FUNCTION_BLOCK FB_ConveyorBase IMPLEMENTS I_Conveyor
VAR_OUTPUT
    initCount : DINT;
    cycleCount : DINT;
END_VAR
VAR
    startup : TON;
    productEdge : R_TRIG;
    delay : TIME;
    requested : BOOL;
    runningState : BOOL;
    lastBlocked : BOOL;
    alarmText : STRING(80);
    count : DINT;
    speed : REAL;
END_VAR

(* All behavior is called through the interface methods. *)

METHOD PUBLIC FB_init : BOOL
VAR_INPUT
    bInitRetains : BOOL;
    bInCopyCode : BOOL;
    startDelay : TIME;
END_VAR
delay := startDelay;
initCount := initCount + 1;
FB_init := TRUE;
END_METHOD

METHOD PUBLIC Start
IF alarmText = '' THEN requested := TRUE; END_IF;
END_METHOD

METHOD PUBLIC Stop
requested := FALSE;
runningState := FALSE;
startup(IN := FALSE, PT := delay);
END_METHOD

METHOD PUBLIC Reset
IF NOT lastBlocked THEN alarmText := ''; END_IF;
END_METHOD

METHOD PROTECTED DetectJam : BOOL
VAR_INPUT
    blocked : BOOL;
END_VAR
DetectJam := FALSE;
END_METHOD

METHOD PUBLIC Cycle
VAR_INPUT
    enabled : BOOL;
    sensor : BOOL;
    blocked : BOOL;
END_VAR
cycleCount := cycleCount + 1;
lastBlocked := blocked;
IF THIS^.DetectJam(blocked := blocked) THEN
    alarmText := 'Jammed';
    requested := FALSE;
END_IF;
startup(IN := requested AND enabled AND alarmText = '', PT := delay);
runningState := startup.Q;
productEdge(CLK := sensor);
IF runningState AND productEdge.Q THEN count := count + 1; END_IF;
END_METHOD

PROPERTY PUBLIC Running : BOOL
GET
Running := runningState;
END_GET
END_PROPERTY

PROPERTY PUBLIC Alarm : STRING(80)
GET
Alarm := alarmText;
END_GET
END_PROPERTY

PROPERTY PUBLIC ProductCount : DINT
GET
ProductCount := count;
END_GET
END_PROPERTY

PROPERTY PUBLIC ActualSpeed : REAL
GET
IF runningState THEN ActualSpeed := speed; ELSE ActualSpeed := 0.0; END_IF;
END_GET
END_PROPERTY

PROPERTY PUBLIC SpeedSetpoint : REAL
GET
SpeedSetpoint := speed;
END_GET
SET
speed := SpeedSetpoint;
END_SET
END_PROPERTY

END_FUNCTION_BLOCK

(* stored: Version 1.1.0.1, ProductVersion 3.1 *)
